(* PLC project Vn_fn_left, Beckhoff Automation GmbH TwinCAT PLC Control 3.5.13.21 *)
(* stored: creationDateTime 1970-01-01T00:00:00 *)

PROGRAM Vn_fn_left

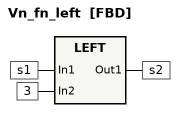
(* FBD diagram, written out as Structured Text *)
s2 := LEFT(s1, 3);
END_PROGRAM
